(* IEC 61131-3 sources: Jacob-Formschaumtechnik-ISEL-CNC-Retrofit/twincat/PLC/src/0_Main, 9 files *)

(* ---- GVL_AlarmCatalog.st ---- *)
(* Meldekatalog, einzige Quelle fuer ID und Klasse je Slot (Befund 11). Slot-Nummer = Index in aCond,
   siehe E_AlarmSlot. Klassen: 0 Info, 1 Warnung, 2 Vorschubhalt, 3 Abbruch, 4 Antriebe aus.
   Slot 12 (Referenzverlust) ist R1, Slot 13 (HMI-Verbindung) R2. Texte pflegt die HMI-Seite. *)
VAR_GLOBAL CONSTANT
    aAlarmId    : ARRAY[0..14] OF INT := [100, 101, 110, 120, 200, 201, 202, 203, 300, 301, 302, 310, 320, 330, 900];
    (* Befund 15: 200 (FU-Stoerung) und 302 (Endschalter) sind R3 statt R4. Die Achsregler bleiben an,
       das Programm wird abgebrochen, vom Endschalter kann in Hand freigefahren werden. [Annahme, mit Kunde abstimmen] *)
    aAlarmClass : ARRAY[0..14] OF INT := [4, 3, 3, 2, 3, 3, 3, 1, 4, 4, 3, 4, 1, 2, 4];
END_VAR

(* ---- GVL_Config.st ---- *)
(* Build-Konfiguration (Befund 9). Die Antriebsabbildung wird hier gewaehlt. Solange nur das
   Simulationsabbild fertig ist, laeuft die Maschine nur damit. Fuer jede andere Variante bleibt die
   Maschine gesperrt (FB_AxisMap_Canopen meldet Fehler FFFF0001), bis die echte Abbildung existiert.
   Auf einer realen Maschine darf bSimulationBuild nicht TRUE sein. *)
VAR_GLOBAL CONSTANT
    eDriveVariant   : E_DriveVariant := E_DriveVariant.Simulation;
    bSimulationBuild: BOOL := (eDriveVariant = E_DriveVariant.Simulation);   (* G-06: nie getrennt von der Antriebsvariante setzen *)
    sSwVersion      : STRING(15) := '0.12.0';   (* G-18: bei jedem Tag mitpflegen, auch in FB_ParamInit *)
    (* Befund 20: Maschinenkennung kommt aus GVL_Persistent.nMachineId, nicht aus dem Code.
       Nur im Simulationsbuild gilt bei nicht gesetzter Kennung (0) die Kennung 1 [Annahme]. *)
    nMachineIdSimDefault : UINT := 1;
    (* Achsnummerierung zentral (Befund 16). HMI- und CNC-Achse: 1 = X, 2 = Y, 3 = Z [Annahme CNC-Kanal].
       Referenzgruppe: 1 = Z, 2 = X, 3 = Y. Antrieb: 1 = Y1, 2 = Y2, 3 = X, 4 = Z [Annahme]. *)
    aHmiAxisToGroup  : ARRAY[1..3] OF USINT := [2, 3, 1];
    aGroupToHmiAxis  : ARRAY[1..3] OF USINT := [3, 1, 2];
    aDriveToHmiAxis  : ARRAY[1..4] OF USINT := [2, 2, 1, 3];
    aDriveToGroup    : ARRAY[1..4] OF USINT := [3, 3, 2, 1];
    (* Befund 15: Verzoegerung der Reglerabschaltung bei R4, damit die CNC gefuehrt bremst [Annahme] *)
    tR4DriveOffDelay : TIME := T#500MS;
END_VAR

(* ---- GVL_HMI.st ---- *)
VAR_GLOBAL
    stCmd : ST_HmiCmd;     (* HMI -> SPS *)
    stSts : ST_HmiSts;     (* SPS -> HMI *)
    stJournal : ST_HmiJournal;  (* SPS -> HMI, Meldejournal (Befund 21), Kopie von GVL_Persistent.stJournal *)
END_VAR

(* ---- GVL_HmiCnc.st ---- *)
VAR_GLOBAL
    stCncSts : ST_HmiCncSts;     (* SPS -> HMI *)
    stCncCmd : ST_HmiCncCmd;     (* HMI -> SPS *)
END_VAR

(* ---- GVL_IO.st ---- *)
(* Prozessabbild der Maschine. Die Verknuepfung mit den Klemmen erfolgt erst nach
   Klemmenwahl und Schaltplan, bis dahin gibt es hier nur Variablen ohne Adresse (Simulation).
   Ruhestrom: FALSE = Fehler/ausgeloest bei allen Sicherheits- und Endschaltersignalen. *)
VAR_GLOBAL
    (* Eingaenge *)
    bSafetyRelayFeedback : BOOL;   (* Pilz-Relais Rueckmeldung *)
    bDoorClosed          : BOOL;
    bAirOk               : BOOL;
    bExtractionOk        : BOOL;
    bFuReady             : BOOL;   (* Commander SK bereit *)
    bFuAtSpeed           : BOOL;   (* [Annahme] Drehzahl erreicht *)
    bSpindlePtcOk        : BOOL;
    bKeyAuto             : BOOL;   (* [offen] nur falls Schluesselschalter vorhanden *)
    bFieldbusOk          : BOOL;   (* EtherCAT/CANopen Status *)
    (* Ausgaenge *)
    bSpindleRun          : BOOL;
    bSpindleCcw          : BOOL;
    rSpindleVolt         : REAL;   (* EL4002 Kanal 1, 0..10 V *)
    bExtractionOut       : BOOL;
    bBlowAirOut          : BOOL;
    bVacuumOut           : BOOL;
    (* Achsen, vier Stueck: 1=Y1 Portal links, 2=Y2 Portal rechts, 3=X Quer, 4=Z [Annahme] *)
    aAxis                : ARRAY[1..4] OF ST_AxisDrive;
    (* Einspeisung fuer Simulation und Test (wirkt nur im Simulationsabbild FB_AxisMap_Simulation) *)
    aSimLimitPlus  : ARRAY[1..4] OF BOOL;
    aSimLimitMinus : ARRAY[1..4] OF BOOL;
    aSimFault      : ARRAY[1..4] OF BOOL;
END_VAR

(* ---- GVL_Machine.st ---- *)
(* Zustandsgroessen und CNC-Schnittstelle (Signale aus/zur CNC kommen spaeter ueber Tc2_CncHli). *)
VAR_GLOBAL
    stParams       : ST_MachineParams;
    bParamsLoaded  : BOOL;
    (* von der CNC [offen, HLI-Anbindung folgt] *)
    nCncMCode      : INT;
    bCncMStrobe    : BOOL;
    nCncToolNo     : UINT;
    bCncProgramDone: BOOL;
    bCncProgramActive : BOOL;  (* Programm laeuft oder Achsen fahren noch (Befund 4) *)
    rCncSpindleRpm : REAL;     (* S-Wert aus dem NC-Programm, 1/min (Befund 10) *)
    aCncHomed      : ARRAY[1..3] OF BOOL;
    (* zur CNC *)
    bCncStartReq   : BOOL;
    bCncHoldReq    : BOOL;
    bCncAbortReq   : BOOL;
    bCncMAck       : BOOL;
    bCncJogPlus    : BOOL;
    bCncJogMinus   : BOOL;
    nCncJogAxis    : USINT;
    bCncJogRapid   : BOOL;
    bCncHomeReq    : BOOL;
    nCncHomeGroup  : USINT;
    bCncSingleBlock: BOOL;
    bCncDryRun     : BOOL;
    bCncOptStop    : BOOL;
    rCncJogStepMm  : REAL;
    bCncHandwheel  : BOOL;
    nCncHandwheelAxis  : USINT;
    nCncHandwheelRatio : USINT;
    bHasHandwheel  : BOOL;     (* [offen] nur M1 mit Bestandsgeraet *)
    bCncJogCreep   : BOOL;     (* Freifahren vom Endschalter: CNC soll im Schleichgang tippen (HLI-Anbindung offen) *)
END_VAR

(* ---- GVL_Persistent.st ---- *)
{attribute 'qualified_only'}
(* Persistente Daten (Befunde 20 und 21). Ueberleben Neustart und Online-Change.
   nMachineId ist die Maschinenkennung des Geraets, gesetzt bei der Inbetriebnahme (0 = nicht gesetzt,
   Maschine bleibt gesperrt, Meldung 900). Damit laeuft ein Softwarestand auf allen Maschinen (LH-2.11.4).
   [offen] Schreibweg ueber die Service-Seite der HMI, bis dahin per ADS. *)
VAR_GLOBAL PERSISTENT
    nMachineId    : UINT;
    nOperatingSec : UDINT;            (* Betriebssekunden *)
    nSpindleSec   : UDINT;            (* Spindellaufzeit in Sekunden *)
    stJournal     : ST_HmiJournal;    (* Meldejournal *)
END_VAR

(* ---- PRG_Main.st ---- *)
(* Hauptprogramm. Aufrufreihenfolge fest: Eingaenge -> Sicherheit -> Achsen -> Meldungen ->
   Verriegelungen -> Zustand -> Geraete -> HMI-Status. Rueckwirkungen zwischen den Bausteinen
   laufen bewusst mit einem Zyklus Verzoegerung, damit keine Schleifen entstehen. *)
PROGRAM PRG_Main
VAR
    fbParamInit: FB_ParamInit;
    fbCncMirror: FB_CncMirror;
    fbParam    : FB_ParamCheck;
    aGrpOfAxis : ARRAY[1..4] OF INT := [3, 3, 2, 1];   (* Achse 1,2 (Y1,Y2) = Gruppe 3, Achse 3 (X) = Gruppe 2, Achse 4 (Z) = Gruppe 1 *)
    fbSafety   : FB_SafetyMonitor;
    fbAxisSim  : ARRAY[1..4] OF FB_AxisMap_Simulation;
    fbSupervisor : FB_AxisSupervisor;
    fbAlarms   : FB_AlarmList;
    fbJournal  : FB_AlarmJournal;
    fbInterlocks : FB_Interlocks;
    fbState    : FB_MachineState;
    fbMode     : FB_OpModeManager;
    fbSpindle  : FB_Spindle;
    fbMFunc    : FB_MFunctions;
    fbTool     : FB_ToolChange;
    fbHoming   : FB_Homing;
    fbJog      : FB_Jog;
    aCond      : ARRAY[0..14] OF BOOL;
    aHomeReq   : ARRAY[1..3] OF BOOL;
    fbAxisCan  : ARRAY[1..4] OF FB_AxisMap_Canopen;
    tonExtraction : TON;
    i          : INT;
    bStandstill: BOOL;
    bSimulation: BOOL := TRUE;     (* bis die Hardwareabbildung steht, immer Simulation *)
    nVersionDummy : INT;
    tonUptime  : TON;
    tonSpindleUptime : TON;
    dwSecTick  : UDINT;
    dtNow      : DT;
    nMachineIdEff : UINT;     (* wirksame Maschinenkennung (Befund 20) *)
    nSysTime   : ULINT;       (* UTC, 100 ns seit 1.1.1601 *)
    bLimitFreeRun : BOOL;     (* Freifahren vom Endschalter erlaubt (Befund 15) *)
    bOtherR3   : BOOL;
    nCls       : INT;
    bHandSpindleBlock : BOOL; (* Hand-Spindel gesperrt bis bSpindleOn einmal FALSE war (Lebenszeichen weg, nicht Hand) *)
    bHandSpindleOn : BOOL;    (* wirksame Hand-Anforderung Spindel *)
    tofModeBlocked : TOF;     (* Hinweis "Betriebsartwechsel abgelehnt" fuer die HMI halten *)
    bLimHitPlus      : BOOL;
    bLimHitMinus     : BOOL;
    bJogPlusBlocked  : BOOL;
    bJogMinusBlocked : BOOL;
    rtHandOn         : R_TRIG;
    bHandCcw         : BOOL;
    bDryRunEff       : BOOL;
    bSpindleLocked   : BOOL;
    bVacuumReq       : BOOL;
    bHomingLostInRun : BOOL;
    bToolChangeDoor  : BOOL;
END_VAR

(* 1. Parameter: initialisieren und pruefen, bei unplausiblen Werten bleibt die Maschine gesperrt *)
(* Befund 20: Kennung aus dem Geraet (persistent), nur im Simulationsbuild Ersatzwert bei 0 *)
nMachineIdEff := GVL_Persistent.nMachineId;
IF nMachineIdEff = 0 AND GVL_Config.bSimulationBuild THEN nMachineIdEff := GVL_Config.nMachineIdSimDefault; END_IF
fbParamInit(nMachineId := nMachineIdEff, stParams := GVL_Machine.stParams);
GVL_Machine.bParamsLoaded := fbParamInit.bLoaded;
fbParam(nIdExpected := nMachineIdEff, nIdLoaded := GVL_Machine.stParams.nMachineId,
        sVerExpected := GVL_Machine.stParams.sSwVersionExpected, sVerRunning := GVL_Config.sSwVersion,
        bParamsLoaded := GVL_Machine.bParamsLoaded);

(* 2. Sicherheit *)
fbSafety(bRelayFeedbackOk := GVL_IO.bSafetyRelayFeedback, bDoorClosed := GVL_IO.bDoorClosed,
         bFieldbusOk := GVL_IO.bFieldbusOk, bAck := GVL_HMI.stCmd.bAck, bAirOk := GVL_IO.bAirOk);

(* 3. Achsen *)
FOR i := 1 TO 4 DO
    GVL_IO.aAxis[i].bEnableReq := fbState.bEnableDrives;
    GVL_IO.aAxis[i].bResetReq  := GVL_HMI.stCmd.bAck;     (* Antriebsfehler quittieren (Befund 14) *)
    IF GVL_Config.eDriveVariant = E_DriveVariant.Simulation THEN
    fbAxisSim[i](bSafeEnable := fbSafety.bDrivesAllowed,
                 bHomeReset := fbHoming.aResetHomed[GVL_Config.aDriveToGroup[i]],
                 bHomeCmd := fbHoming.bHomeCmd AND fbHoming.nActiveGroup = GVL_Config.aDriveToGroup[i],
                 bInjLimitPlus := GVL_IO.aSimLimitPlus[i], bInjLimitMinus := GVL_IO.aSimLimitMinus[i],
                 bInjFault := GVL_IO.aSimFault[i],
                 stAxis := GVL_IO.aAxis[i]);
    ELSE
        (* Befund 9: echte Abbildung fehlt, FB_AxisMap_Canopen sperrt die Maschine (Fehler FFFF0001) *)
        fbAxisCan[i](bSafeEnable := fbSafety.bDrivesAllowed, stAxis := GVL_IO.aAxis[i]);
    END_IF
END_FOR
(* Einheitlicher Referenzstatus (Befund 3): einzige Quelle ist GVL_IO.aAxis[].bHomed.
   Gruppen 1 = Z, 2 = X, 3 = Y (beide Portalseiten). *)
GVL_Machine.aCncHomed[1] := GVL_IO.aAxis[4].bHomed;
GVL_Machine.aCncHomed[2] := GVL_IO.aAxis[3].bHomed;
GVL_Machine.aCncHomed[3] := GVL_IO.aAxis[1].bHomed AND GVL_IO.aAxis[2].bHomed;
GVL_HmiCnc.stCncSts.aAxis[1].bHomed := GVL_Machine.aCncHomed[2];   (* HMI-Achse 1 = X *)
GVL_HmiCnc.stCncSts.aAxis[2].bHomed := GVL_Machine.aCncHomed[3];   (* HMI-Achse 2 = Y *)
GVL_HmiCnc.stCncSts.aAxis[3].bHomed := GVL_Machine.aCncHomed[1];   (* HMI-Achse 3 = Z *)
fbSupervisor(bEnableCmd := fbState.bEnableDrives, bFieldbusOk := GVL_IO.bFieldbusOk,
             bHomingActive := fbHoming.bBusy, rMaxFollowErr := 1.0, aAxis := GVL_IO.aAxis);
bStandstill := fbSpindle.bStandstillOk AND fbState.eState <> E_MachState.Execute AND NOT fbJog.bJogPlusReq AND NOT fbJog.bJogMinusReq;

(* 4. Meldungen *)
(* Werkzeugwechsel mit Tuerfreigabe: Tuer offen und Spindel steht. Dann sind Tuer-Meldung und das dadurch abfallende
   Sicherheitsrelais kein Abbruchgrund, das Programm bleibt gehalten. Sonst ist eine offene Tuer weiter ein Abbruch. *)
bToolChangeDoor := fbTool.bDoorRelease AND NOT GVL_IO.bDoorClosed AND GVL_IO.bFieldbusOk;
aCond[0]  := NOT GVL_IO.bSafetyRelayFeedback AND NOT bToolChangeDoor;
aCond[1]  := NOT GVL_IO.bDoorClosed AND NOT bToolChangeDoor;
aCond[2]  := GVL_Machine.stParams.bAirMonitoring AND NOT GVL_IO.bAirOk;
(* Absaugung: Rueckmeldung darf nach dem Einschalten tFeedbackTimeout dauern (Befund 12) *)
tonExtraction(IN := NOT GVL_IO.bExtractionOk AND GVL_IO.bExtractionOut, PT := GVL_Machine.stParams.tFeedbackTimeout);
aCond[3]  := tonExtraction.Q;
aCond[4]  := NOT GVL_IO.bFuReady;
aCond[5]  := fbSpindle.bPtcTrip;
aCond[6]  := fbSpindle.bNoFeedback;
aCond[7]  := fbSpindle.bLockedSetup;
aCond[8]  := fbSupervisor.bAnyFault OR fbSupervisor.bEnableTimeout;
aCond[9]  := fbSupervisor.bFollowErr;
aCond[10] := fbSupervisor.bAnyHwLimit;
aCond[11] := NOT GVL_IO.bFieldbusOk;
aCond[12] := fbSupervisor.bHomingLost;
aCond[13] := NOT fbJog.bHmiLinkOk;
aCond[14] := fbParam.bMismatch;
fbAlarms(aCond := aCond, bAck := GVL_HMI.stCmd.bAck);
(* Befund 21: Zeitstempel UTC, Journal persistent, HMI liest die Kopie *)
nSysTime := F_GetSystemTime();
IF nSysTime > 116444736000000000 THEN
    dtNow := DWORD_TO_DT(ULINT_TO_DWORD((nSysTime - 116444736000000000) / 10000000));
END_IF
fbJournal(aCond := aCond, aId := GVL_AlarmCatalog.aAlarmId, aClass := GVL_AlarmCatalog.aAlarmClass,
          dtNow := dtNow, stJournal := GVL_Persistent.stJournal);
GVL_HMI.stJournal := GVL_Persistent.stJournal;

(* Befund 15: Steht nur der Endschalter (302, R3) an, darf in Hand im Schleichgang freigefahren werden.
   [offen] Richtungssperre zur Endschalterseite liegt in CNC/Antrieb (Softwareendlage, Endschalterlogik). *)
bOtherR3 := FALSE;
FOR i := 0 TO 14 DO
    nCls := GVL_AlarmCatalog.aAlarmClass[i];
    IF i <> 10 (* E_AlarmSlot.HwLimitHit *) AND nCls >= 3 AND (fbAlarms.aList[i].bActive OR fbAlarms.aList[i].bLatched) THEN
        bOtherR3 := TRUE;
    END_IF
END_FOR
bLimitFreeRun := aCond[10] AND NOT bOtherR3;   (* Slot 10 = E_AlarmSlot.HwLimitHit *)

(* 5. Betriebsart und Verriegelungen *)
(* Befund 17: Wechsel nur im echten Stillstand, ohne Referenzfahrt und ohne offene Werkzeugwechsel-Aufforderung *)
fbMode(eRequest := GVL_HMI.stCmd.eModeRequest,
       bStandstill := bStandstill AND fbInterlocks.bModeChangeOk AND NOT fbHoming.bBusy AND NOT fbTool.bRequest,
       bHasKeySwitch := FALSE, bKeyAuto := GVL_IO.bKeyAuto);
(* Abgelehnter Wunsch wird verworfen, sonst fuehrte die SPS ihn beim naechsten Stillstand verspaetet aus.
   Der Hinweis bleibt 3 s fuer die HMI stehen. *)
IF fbMode.bChangeBlocked THEN
    GVL_HMI.stCmd.eModeRequest := fbMode.eMode;
END_IF
tofModeBlocked(IN := fbMode.bChangeBlocked, PT := T#3S);
fbInterlocks(eMode := fbMode.eMode, eState := fbState.eState, bSafetyOk := fbSafety.bSafetyOk,
             bAllHomed := fbSupervisor.bAllHomed, bDrivesEnabled := fbSupervisor.bAllEnabled,
             bHmiLinkOk := fbJog.bHmiLinkOk, bAnyR2OrHigher := fbAlarms.bAnyR2OrHigher,
             bAnyR3OrHigher := fbAlarms.bAnyR3OrHigher, bAirOk := GVL_IO.bAirOk OR NOT GVL_Machine.stParams.bAirMonitoring,
             bHomingBusy := fbHoming.bBusy, bLimitFreeRun := bLimitFreeRun);

(* 6. Zustand *)
(* G-10: Geht die Referenz im laufenden oder gehaltenen Programm verloren, wirkt das wie R3 (Abbruch). Sonst nur Warnung R1. *)
bHomingLostInRun := fbSupervisor.bHomingLost AND (fbState.eState = E_MachState.Execute OR fbState.eState = E_MachState.Held);
fbState(bSafetyOk := fbSafety.bSafetyOk, bDrivesAllowed := fbSafety.bDrivesAllowed,
        bAnyR2OrHigher := fbAlarms.bAnyR2OrHigher OR bHomingLostInRun,
        bAnyR3OrHigher := fbAlarms.bAnyR3OrHigher OR bHomingLostInRun,
        bAnyR4 := fbAlarms.bAnyR4, bAckPending := fbAlarms.bAckPending,
        bStartOk := fbInterlocks.bProgramStartOk AND NOT fbTool.bHoldProgram,
        bStartCmd := GVL_HMI.stCmd.bStart, bHoldCmd := GVL_HMI.stCmd.bHold OR fbMFunc.bProgramHalt,
        bAbortCmd := GVL_HMI.stCmd.bAbort, bProgramDone := GVL_Machine.bCncProgramDone,
        bProgramActive := GVL_Machine.bCncProgramActive,
        bAck := GVL_HMI.stCmd.bAck, tR4OffDelay := GVL_Config.tR4DriveOffDelay,
        bDoorOpenAllowed := bToolChangeDoor);

(* 7. Geraete: Spindel (M3/M4 aus Programm, in Hand von der HMI) *)
(* Hand-Spindel: Nach Lebenszeichenverlust oder ausserhalb Hand setzt die SPS bSpindleOn zurueck und sperrt,
   bis bSpindleOn FALSE gesehen wurde. Ein stehender Pegel startet die Spindel so nie von selbst wieder. *)
IF NOT fbJog.bHmiLinkOk OR fbMode.eMode <> E_OpMode.Hand THEN
    bHandSpindleBlock := TRUE;
    GVL_HMI.stCmd.bSpindleOn := FALSE;
ELSIF NOT GVL_HMI.stCmd.bSpindleOn THEN
    bHandSpindleBlock := FALSE;
END_IF
bHandSpindleOn := GVL_HMI.stCmd.bSpindleOn AND NOT bHandSpindleBlock;
(* G-11: Drehrichtung wird beim Einschalten festgehalten, Umschalten bei laufender oder wartender Spindel startet nichts *)
rtHandOn(CLK := bHandSpindleOn);
IF rtHandOn.Q THEN bHandCcw := GVL_HMI.stCmd.bSpindleCcw; END_IF
(* G-12: Trockenlauf wirkt nur in Auto und nur so, wie er beim Programmstart stand (nicht mitten im Programm) *)
IF fbState.eState <> E_MachState.Execute AND fbState.eState <> E_MachState.Held THEN
    bDryRunEff := GVL_HMI.stCmd.bDryRun;
END_IF
bSpindleLocked := fbMode.eMode = E_OpMode.Setup OR (fbMode.eMode = E_OpMode.Auto AND bDryRunEff);
fbMFunc(nMCode := GVL_Machine.nCncMCode, bMStrobe := GVL_Machine.bCncMStrobe,
        bSpindleOk := fbInterlocks.bSpindleOk, bAuxOk := fbInterlocks.bAuxOk,
        bReset := fbState.bSpindleStop OR GVL_Machine.bCncProgramDone, bOptStop := GVL_HMI.stCmd.bOptStop,
        bSpindleRunning := fbSpindle.bRunning, bSpindleSkip := bSpindleLocked);
fbSpindle(bRelease := fbInterlocks.bSpindleOk AND NOT fbState.bSpindleStop AND NOT fbTool.bSpindleLock,
          bStop := fbState.bSpindleStop,
          bSetupLocked := bSpindleLocked,
          bAllowPend := fbMode.eMode = E_OpMode.Auto,   (* G-11: nur das Programm darf auf Stillstand warten, Hand-Start wird sonst verworfen *)
          bStartCw := (fbMFunc.bSpindleCw AND fbMode.eMode = E_OpMode.Auto) OR (bHandSpindleOn AND NOT bHandCcw),
          bStartCcw := (fbMFunc.bSpindleCcw AND fbMode.eMode = E_OpMode.Auto) OR (bHandSpindleOn AND bHandCcw),
          rSetRpm := SEL(fbMode.eMode = E_OpMode.Auto, GVL_HMI.stCmd.rSpindleSetRpm, GVL_Machine.rCncSpindleRpm),
          rOverridePct := UINT_TO_REAL(GVL_HmiCnc.stCncSts.nOvrSpindle),
          bFuReady := GVL_IO.bFuReady, bFuAtSpeed := GVL_IO.bFuAtSpeed, bPtcOk := GVL_IO.bSpindlePtcOk,
          bAckReset := GVL_HMI.stCmd.bAck, rMaxRpm := GVL_Machine.stParams.rSpindleMaxRpm,
          rMinRpm := GVL_Machine.stParams.rSpindleMinRpm, rVoltMax := GVL_Machine.stParams.rSpindleVoltMax,
          tRunUp := GVL_Machine.stParams.tSpindleRunUp, tStandstill := GVL_Machine.stParams.tSpindleStandstill);
GVL_IO.bSpindleRun  := fbSpindle.bRunCmd;
GVL_IO.bSpindleCcw  := fbSpindle.bDirCcw;
GVL_IO.rSpindleVolt := fbSpindle.rVoltOut;

fbTool(bM6Request := fbMFunc.bToolChangeReq, nToolNo := GVL_Machine.nCncToolNo,
       bSpindleStopped := fbSpindle.bStandstillOk, bConfirm := GVL_HMI.stCmd.bToolChangeDone,
       bAbort := GVL_HMI.stCmd.bAbort OR fbState.eState = E_MachState.EStop OR fbState.eState = E_MachState.Aborted
                 OR fbState.eState = E_MachState.Fault);   (* G-05: Anforderung faellt bei Abbruch, R3 und NOT-HALT *)

(* Hilfsausgaenge: von Hand oder per M-Code, nur mit Freigabe *)
GVL_IO.bExtractionOut := fbInterlocks.bAuxOk AND (fbMFunc.bExtraction OR GVL_HMI.stCmd.bExtraction);
GVL_IO.bBlowAirOut    := fbInterlocks.bAuxOk AND (fbMFunc.bBlowAir OR GVL_HMI.stCmd.bBlowAir);
(* G-04: Vakuum (Werkstueckspannung) bleibt bei Abbruch und NOT-HALT gehalten. Einschalten nur mit Freigabe. *)
bVacuumReq := fbMFunc.bVacuum OR GVL_HMI.stCmd.bVacuum;
GVL_IO.bVacuumOut     := bVacuumReq AND (fbInterlocks.bAuxOk OR GVL_IO.bVacuumOut);

(* 8. Referenzieren und Tippen *)
(* Zuordnung HMI-Achse (1=X, 2=Y, 3=Z) zu Referenzgruppe (1=Z, 2=X, 3=Y) *)
aHomeReq[1] := GVL_HMI.stCmd.bHomeAxis[3];
aHomeReq[2] := GVL_HMI.stCmd.bHomeAxis[1];
aHomeReq[3] := GVL_HMI.stCmd.bHomeAxis[2];
fbHoming(bStart := GVL_HMI.stCmd.bHomeRequest, aStartAxis := aHomeReq,
         bAbort := GVL_HMI.stCmd.bAbort OR GVL_HMI.stCmd.bHomeAbort,
         bHomingOk := fbInterlocks.bHomingOk, aHomed := GVL_Machine.aCncHomed);
(* G-01: Endschalter je Seite der gewaehlten Achse (HMI 1=X -> Antrieb 3, 2=Y -> Antriebe 1 und 2, 3=Z -> Antrieb 4).
   Ruhestrom: FALSE = ausgeloest. [Annahme] Tippen+ faehrt zur Plus-Seite. Ist ein Endschalter ausgeloest, ist Tippen
   nur fuer die betroffene Achse und nur in Gegenrichtung erlaubt, ohne Eilgang. *)
bLimHitPlus := FALSE; bLimHitMinus := FALSE;
CASE GVL_HMI.stCmd.nJogAxis OF
    1: bLimHitPlus  := NOT GVL_IO.aAxis[3].bHwLimitPlus;
       bLimHitMinus := NOT GVL_IO.aAxis[3].bHwLimitMinus;
    2: bLimHitPlus  := NOT GVL_IO.aAxis[1].bHwLimitPlus  OR NOT GVL_IO.aAxis[2].bHwLimitPlus;
       bLimHitMinus := NOT GVL_IO.aAxis[1].bHwLimitMinus OR NOT GVL_IO.aAxis[2].bHwLimitMinus;
    3: bLimHitPlus  := NOT GVL_IO.aAxis[4].bHwLimitPlus;
       bLimHitMinus := NOT GVL_IO.aAxis[4].bHwLimitMinus;
END_CASE
bJogPlusBlocked  := bLimHitPlus;
bJogMinusBlocked := bLimHitMinus;
IF aCond[10] AND NOT (bLimHitPlus OR bLimHitMinus) THEN
    bJogPlusBlocked := TRUE; bJogMinusBlocked := TRUE;   (* Endschalter an einer anderen Achse: diese Achse bleibt stehen *)
END_IF
GVL_Machine.bCncJogCreep := bLimitFreeRun;   (* CNC: Freifahren nur im Schleichgang (HLI-Anbindung offen) *)
fbJog(bJogOk := fbInterlocks.bJogOk, bPlus := GVL_HMI.stCmd.bJogPlus, bMinus := GVL_HMI.stCmd.bJogMinus,
      bPlusBlocked := bJogPlusBlocked, bMinusBlocked := bJogMinusBlocked,
      nAxis := GVL_HMI.stCmd.nJogAxis, bRapid := GVL_HMI.stCmd.bJogRapid AND NOT bLimitFreeRun AND GVL_HmiCnc.stCncSts.nSpeedLimitActivePct >= 50,
      nHeartbeat := GVL_HMI.stCmd.nHeartbeat, tHmiTimeout := GVL_Machine.stParams.tHmiTimeout);

(* CNC-Spiegel (Simulation, bis TF5200 verfuegbar ist) *)
fbCncMirror(bStandstill := fbState.eState <> E_MachState.Execute AND fbState.eState <> E_MachState.Held
                           AND NOT GVL_Machine.bCncProgramActive,
            stCmd := GVL_HmiCnc.stCncCmd, stSts := GVL_HmiCnc.stCncSts);

(* 9. Anforderungen an die CNC *)
GVL_Machine.bCncStartReq := fbState.bCncStart;
GVL_Machine.bCncHoldReq  := fbState.bCncHold OR fbTool.bHoldProgram;
GVL_Machine.bCncAbortReq := fbState.bCncAbort;
GVL_Machine.bCncMAck     := fbMFunc.bAck;
GVL_Machine.bCncJogPlus  := fbJog.bJogPlusReq;
GVL_Machine.bCncJogMinus := fbJog.bJogMinusReq;
GVL_Machine.nCncJogAxis  := fbJog.nAxisReq;
GVL_Machine.bCncJogRapid := fbJog.bRapidReq;
GVL_Machine.bCncHomeReq  := fbHoming.bHomeCmd;
GVL_Machine.nCncHomeGroup:= fbHoming.nActiveGroup;
GVL_Machine.bCncSingleBlock := GVL_HMI.stCmd.bSingleBlock;
GVL_Machine.bCncDryRun   := bDryRunEff AND fbMode.eMode = E_OpMode.Auto;
GVL_Machine.bCncOptStop  := GVL_HMI.stCmd.bOptStop;
GVL_Machine.rCncJogStepMm := GVL_HMI.stCmd.rJogStepMm;
(* Handrad: nur freigegeben, wenn vorhanden, in Hand und Tippen erlaubt *)
GVL_Machine.bCncHandwheel := GVL_Machine.bHasHandwheel AND GVL_HMI.stCmd.bHandwheelEnable AND fbInterlocks.bJogOk;
GVL_Machine.nCncHandwheelAxis  := GVL_HMI.stCmd.nHandwheelAxis;
GVL_Machine.nCncHandwheelRatio := GVL_HMI.stCmd.nHandwheelRatio;

(* 10. Status an die HMI *)
(* Befund 21: Betriebs- und Spindellaufzeit persistent, Sekundentakt *)
tonUptime(IN := TRUE, PT := T#1S);
IF tonUptime.Q THEN
    dwSecTick := dwSecTick + 1;
    GVL_Persistent.nOperatingSec := GVL_Persistent.nOperatingSec + 1;
    IF fbSpindle.bRunCmd THEN GVL_Persistent.nSpindleSec := GVL_Persistent.nSpindleSec + 1; END_IF
    tonUptime(IN := FALSE);
END_IF
GVL_HMI.stSts.eMode          := fbMode.eMode;
GVL_HMI.stSts.eState         := fbState.eState;
GVL_HMI.stSts.bSafetyOk      := fbSafety.bSafetyOk;
GVL_HMI.stSts.bDrivesEnabled := fbSupervisor.bAllEnabled;
GVL_HMI.stSts.bAllHomed      := fbSupervisor.bAllHomed;
GVL_HMI.stSts.bHmiLinkOk     := fbJog.bHmiLinkOk;
GVL_HMI.stSts.bSpindleRunning:= fbSpindle.bRunning;
GVL_HMI.stSts.rSpindleActRpm := SEL(fbSpindle.bRunning, 0.0, fbSpindle.rActRpm);   (* Sollwert nur bei Drehzahl erreicht anzeigen (Befund 13) *)
GVL_HMI.stSts.bExtractionOn  := GVL_IO.bExtractionOut;
GVL_HMI.stSts.bBlowAirOn     := GVL_IO.bBlowAirOut;
GVL_HMI.stSts.bVacuumOn      := GVL_IO.bVacuumOut;
GVL_HMI.stSts.bToolChangeReq := fbTool.bRequest;
GVL_HMI.stSts.nToolChangeNo  := fbTool.nRequestedTool;
GVL_HMI.stSts.nTopAlarmId    := fbAlarms.nTopId;
GVL_HMI.stSts.eTopAlarmClass := F_ToFaultClass(fbAlarms.nTopClass);
GVL_HMI.stSts.nActiveAlarms  := fbAlarms.nActive;
GVL_HMI.stSts.nMachineId     := GVL_Machine.stParams.nMachineId;
GVL_HMI.stSts.sSwVersion     := GVL_Config.sSwVersion;
GVL_HMI.stSts.bSimulationActive := GVL_Config.bSimulationBuild;
GVL_HMI.stSts.bModeChangeBlocked := tofModeBlocked.Q;
GVL_HMI.stSts.dwOperatingSec := GVL_Persistent.nOperatingSec;
GVL_HMI.stSts.dwSpindleSec   := GVL_Persistent.nSpindleSec;
GVL_HMI.stSts.nHeartbeatEcho := GVL_HMI.stCmd.nHeartbeat;
GVL_HMI.stSts.bLimitFreeRun  := bLimitFreeRun;
GVL_HMI.stSts.bToolChangeDoorRelease := fbTool.bDoorRelease;
GVL_HMI.stSts.bHandwheelActive := GVL_Machine.bCncHandwheel;
GVL_HMI.stSts.eHomeState[1]  := fbHoming.eHomeState[2];   (* X *)
GVL_HMI.stSts.eHomeState[2]  := fbHoming.eHomeState[3];   (* Y *)
GVL_HMI.stSts.eHomeState[3]  := fbHoming.eHomeState[1];   (* Z *)
GVL_HMI.stSts.nHomeStep      := fbHoming.nStepOut;
GVL_HMI.stSts.aAlarms        := fbAlarms.aList;
GVL_HMI.stSts.aDrive         := GVL_IO.aAxis;
GVL_HMI.stSts.bFieldbusOk    := GVL_IO.bFieldbusOk;
GVL_HMI.stSts.bFuFault       := NOT GVL_IO.bFuReady;
GVL_HMI.stSts.bPtcTrip       := fbSpindle.bPtcTrip;

(* 11. Befund 16: Impulse aus der HMI loescht die SPS nach der Auswertung in diesem Zyklus.
   Die HMI setzt nur TRUE (Einzelfeld schreiben, nicht die ganze Struktur), ein Impuls geht so nie verloren. *)
GVL_HMI.stCmd.bStart          := FALSE;
GVL_HMI.stCmd.bHold           := FALSE;
GVL_HMI.stCmd.bAbort          := FALSE;
GVL_HMI.stCmd.bAck            := FALSE;
GVL_HMI.stCmd.bHomeRequest    := FALSE;
GVL_HMI.stCmd.bHomeAbort      := FALSE;
GVL_HMI.stCmd.bToolChangeDone := FALSE;
GVL_HMI.stCmd.bHomeAxis[1]    := FALSE;
GVL_HMI.stCmd.bHomeAxis[2]    := FALSE;
GVL_HMI.stCmd.bHomeAxis[3]    := FALSE;
GVL_HmiCnc.stCncCmd.bProgramLoad   := FALSE;
GVL_HmiCnc.stCncCmd.bTableWrite    := FALSE;
GVL_HmiCnc.stCncCmd.bWcsSetCurrent := FALSE;
END_PROGRAM

(* ---- PRG_Test.st ---- *)
(* Simulationstest der Grundfunktionen (nur im Simulations-Build, GVL_Config.bSimulationBuild).
   Starten: bTestEnable online auf TRUE setzen. Der Test speist Eingaenge und HMI-Kommandos ein und prueft
   Referenz, Tippen, NOT-HALT und Spindel gegen die Fehlerfaelle aus dem Gutachten (kein Selbstanlauf nach
   Quittierung). Ergebnis: bTestDone, nFails, sFirstFail. Rueckgabe in der Runtime lesen. *)
PROGRAM PRG_Test
VAR
    bTestEnable : BOOL;                 (* online auf TRUE setzen *)
    bTestDone   : BOOL;
    nFails      : INT;
    sFirstFail  : STRING(100);
    nStep       : INT;
    tWait       : TIME;
    tonStep     : TON;
    tonHb       : TON;
    bNext       : BOOL;
    bRelay      : BOOL := TRUE;         (* Rueckmeldung Sicherheitsrelais, NOT-HALT = FALSE *)
    bFailNow    : BOOL;
    sMsg        : STRING(100);
    bHbStop     : BOOL;                 (* TRUE = simuliertes Lebenszeichen der HMI ausgefallen *)
    nIdx        : INT;
    bDoor       : BOOL := TRUE;         (* Tuer geschlossen *)
END_VAR

(* G-06: Der Test schreibt Sicherheitseingaenge und darf nur mit dem Simulationsabbild laufen *)
IF NOT (bTestEnable AND GVL_Config.bSimulationBuild AND GVL_Config.eDriveVariant = E_DriveVariant.Simulation) THEN
    bHbStop := FALSE;
    FOR nIdx := 1 TO 4 DO
        GVL_IO.aSimLimitPlus[nIdx] := FALSE;
        GVL_IO.aSimLimitMinus[nIdx] := FALSE;
        GVL_IO.aSimFault[nIdx] := FALSE;
    END_FOR
    IF nStep <> 0 THEN
        (* Test beendet oder abgebrochen: CNC-Stub einmalig zuruecknehmen *)
        GVL_Machine.bCncProgramActive := FALSE; GVL_Machine.bCncMStrobe := FALSE; GVL_Machine.nCncMCode := 0;
        GVL_Machine.rCncSpindleRpm := 0.0;
    END_IF
    nStep := 0;
    RETURN;
END_IF

(* Simulierte HMI: Lebenszeichen alle 100 ms. Simulierter Umrichter: Drehzahl erreicht folgt dem Start. *)
tonHb(IN := NOT tonHb.Q, PT := T#100MS);
IF tonHb.Q AND NOT bHbStop THEN GVL_HMI.stCmd.nHeartbeat := GVL_HMI.stCmd.nHeartbeat + 1; END_IF
GVL_IO.bFuAtSpeed := GVL_IO.bSpindleRun;

(* Simulierte Eingaenge: alles in Ordnung, nur das Sicherheitsrelais steuert der Test *)
GVL_IO.bSafetyRelayFeedback := bRelay AND bDoor;   (* offene Tuer laesst auch das Pilz-Relais abfallen *)
GVL_IO.bDoorClosed   := bDoor;
GVL_IO.bAirOk        := TRUE;
GVL_IO.bExtractionOk := TRUE;
GVL_IO.bFuReady      := TRUE;
GVL_IO.bSpindlePtcOk := TRUE;
GVL_IO.bFieldbusOk   := TRUE;

tonStep(IN := NOT bNext, PT := tWait);
bNext := FALSE;

CASE nStep OF
    0:  (* Start *)
        nFails := 0; sFirstFail := ''; bTestDone := FALSE; bRelay := TRUE;
        GVL_HMI.stCmd.eModeRequest := E_OpMode.Hand;
        nStep := 10; tWait := T#1S; bNext := TRUE;

    10: (* T01 Anlauf: Maschine startet gelatcht, nicht frei *)
        IF tonStep.Q THEN
            (* Eingaenge sind jetzt in Ordnung, aber ohne Quittierung darf die Maschine nicht frei sein (EStop oder Stopped) *)
            IF GVL_HMI.stSts.eState = E_MachState.Idle OR GVL_HMI.stSts.eState = E_MachState.Execute OR GVL_HMI.stSts.bDrivesEnabled THEN sMsg := 'T01 Anlauf ohne Quittierung frei'; bFailNow := TRUE; END_IF
            GVL_HMI.stCmd.bAck := TRUE;
            nStep := 20; tWait := T#1S; bNext := TRUE;
        END_IF

    20: (* T02 Quittierung -> Idle, dann Referenzfahrt anfordern *)
        IF tonStep.Q THEN
            IF GVL_HMI.stSts.eState <> E_MachState.Idle THEN sMsg := 'T02 Quittierung fuehrt nicht nach Idle'; bFailNow := TRUE; END_IF
            GVL_HMI.stCmd.bHomeRequest := TRUE;
            nStep := 30; tWait := T#20S; bNext := TRUE;
        END_IF

    30: (* T03 Referenzfahrt aller Gruppen *)
        IF GVL_HMI.stSts.bAllHomed THEN
            nStep := 40; tWait := T#500MS; bNext := TRUE;
        ELSIF tonStep.Q THEN
            sMsg := 'T03 Referenzfahrt: Zeitueberschreitung'; bFailNow := TRUE;
            nStep := 40; tWait := T#500MS; bNext := TRUE;
        END_IF

    40: (* Tippen: Achse waehlen, 300 ms stabil *)
        IF tonStep.Q THEN
            GVL_HMI.stCmd.nJogAxis := 1;
            nStep := 50; tWait := T#300MS; bNext := TRUE;
        END_IF

    50: (* Tippen+ starten *)
        IF tonStep.Q THEN
            GVL_HMI.stCmd.bJogPlus := TRUE;
            nStep := 60; tWait := T#500MS; bNext := TRUE;
        END_IF

    60: (* T04 Tippen+ aktiv, dann loslassen *)
        IF tonStep.Q THEN
            IF NOT GVL_Machine.bCncJogPlus THEN sMsg := 'T04 Tippen+ startet nicht'; bFailNow := TRUE; END_IF
            GVL_HMI.stCmd.bJogPlus := FALSE;
            nStep := 70; tWait := T#300MS; bNext := TRUE;
        END_IF

    70: (* T05 Tippen stoppt beim Loslassen, dann Taste wieder druecken *)
        IF tonStep.Q THEN
            IF GVL_Machine.bCncJogPlus THEN sMsg := 'T05 Tippen stoppt nicht beim Loslassen'; bFailNow := TRUE; END_IF
            GVL_HMI.stCmd.bJogPlus := TRUE;
            nStep := 80; tWait := T#400MS; bNext := TRUE;
        END_IF

    80: (* NOT-HALT bei gehaltener Tippen-Taste *)
        IF tonStep.Q THEN
            bRelay := FALSE;
            nStep := 90; tWait := T#500MS; bNext := TRUE;
        END_IF

    90: (* T07 NOT-HALT erkannt, Tippen aus, Antriebe weg *)
        IF tonStep.Q THEN
            IF GVL_HMI.stSts.eState <> E_MachState.EStop THEN sMsg := 'T07 NOT-HALT nicht erkannt'; bFailNow := TRUE; END_IF
            IF GVL_Machine.bCncJogPlus THEN sMsg := 'T07b Tippen laeuft bei NOT-HALT weiter'; bFailNow := TRUE; END_IF
            IF GVL_HMI.stSts.bDrivesEnabled THEN sMsg := 'T07c Antriebe bleiben bei NOT-HALT frei'; bFailNow := TRUE; END_IF
            bRelay := TRUE;
            nStep := 100; tWait := T#500MS; bNext := TRUE;
        END_IF

    100: (* T08/T06 Sicherheitskreis wieder zu: kein Wiederanlauf, gehaltene Taste startet nichts *)
        IF tonStep.Q THEN
            IF GVL_HMI.stSts.eState <> E_MachState.EStop THEN sMsg := 'T08 NOT-HALT ohne Quittierung verlassen'; bFailNow := TRUE; END_IF
            IF GVL_Machine.bCncJogPlus THEN sMsg := 'T06 Tippen startet nach NOT-HALT von selbst'; bFailNow := TRUE; END_IF
            GVL_HMI.stCmd.bAck := TRUE;
            nStep := 110; tWait := T#1500MS; bNext := TRUE;
        END_IF

    110: (* T09 Quittierung -> Idle, gehaltene Tippen-Taste startet nicht, dann Spindel in Hand *)
        IF tonStep.Q THEN
            IF GVL_HMI.stSts.eState <> E_MachState.Idle THEN sMsg := 'T09 Quittierung nach NOT-HALT fuehrt nicht nach Idle'; bFailNow := TRUE; END_IF
            IF GVL_Machine.bCncJogPlus THEN sMsg := 'T06b Tippen startet nach Quittierung von selbst'; bFailNow := TRUE; END_IF
            GVL_HMI.stCmd.bJogPlus := FALSE;
            GVL_HMI.stCmd.rSpindleSetRpm := 12000.0;
            GVL_HMI.stCmd.bSpindleOn := TRUE;
            nStep := 120; tWait := T#1500MS; bNext := TRUE;
        END_IF

    120: (* T10 Spindel startet in Hand, Spannung passt zur Drehzahl *)
        IF tonStep.Q THEN
            IF NOT GVL_IO.bSpindleRun THEN sMsg := 'T10 Spindel startet nicht (Hand)'; bFailNow := TRUE; END_IF
            IF ABS(GVL_IO.rSpindleVolt - 7.2) > 0.3 THEN sMsg := 'T10b Spindelspannung passt nicht zu 12000 1/min'; bFailNow := TRUE; END_IF
            bRelay := FALSE;
            nStep := 130; tWait := T#400MS; bNext := TRUE;
        END_IF

    130: (* T11 Spindel stoppt bei NOT-HALT *)
        IF tonStep.Q THEN
            IF GVL_IO.bSpindleRun THEN sMsg := 'T11 Spindel laeuft bei NOT-HALT weiter'; bFailNow := TRUE; END_IF
            bRelay := TRUE;
            nStep := 140; tWait := T#500MS; bNext := TRUE;
        END_IF

    140: (* Quittieren, Spindeltaste bleibt gedrueckt *)
        IF tonStep.Q THEN
            GVL_HMI.stCmd.bAck := TRUE;
            nStep := 150; tWait := T#1500MS; bNext := TRUE;
        END_IF

    150: (* T12 kein Selbstanlauf der Spindel nach Quittierung *)
        IF tonStep.Q THEN
            IF GVL_IO.bSpindleRun THEN sMsg := 'T12 Spindel startet nach Quittierung von selbst'; bFailNow := TRUE; END_IF
            GVL_HMI.stCmd.bSpindleOn := FALSE;
            nStep := 160; tWait := T#11S; bNext := TRUE;   (* Auslaufzeit abwarten: Hand-Start waehrend des Auslaufs wird verworfen (G-11) *)
        END_IF

    160: (* Spindel erneut starten (Auslaufzeit abwarten), danach HMI-Verlust *)
        IF tonStep.Q THEN
            GVL_HMI.stCmd.bSpindleOn := TRUE;
            nStep := 170; tWait := T#13S; bNext := TRUE;
        END_IF

    170: (* T13a Spindel laeuft, dann Lebenszeichen der HMI ausfallen lassen *)
        IF tonStep.Q THEN
            IF NOT GVL_IO.bSpindleRun THEN sMsg := 'T13a Spindel startet nach Stillstand nicht'; bFailNow := TRUE; END_IF
            bHbStop := TRUE;
            nStep := 180; tWait := T#1500MS; bNext := TRUE;
        END_IF

    180: (* T13 Spindel stoppt bei HMI-Verlust, Meldung 330 steht *)
        IF tonStep.Q THEN
            IF GVL_IO.bSpindleRun THEN sMsg := 'T13 Spindel laeuft bei HMI-Verlust weiter'; bFailNow := TRUE; END_IF
            IF NOT GVL_HMI.stSts.aAlarms[13].bActive THEN sMsg := 'T13b Meldung 330 (HMI-Verbindung) fehlt'; bFailNow := TRUE; END_IF
            bHbStop := FALSE;
            nStep := 190; tWait := T#1500MS; bNext := TRUE;
        END_IF

    190: (* T14 kein Selbstanlauf der Spindel bei Rueckkehr der HMI *)
        IF tonStep.Q THEN
            IF GVL_IO.bSpindleRun THEN sMsg := 'T14 Spindel startet bei Rueckkehr der HMI von selbst'; bFailNow := TRUE; END_IF
            GVL_HMI.stCmd.bSpindleOn := FALSE;
            nStep := 300; tWait := T#500MS; bNext := TRUE;
        END_IF

    300: (* G-01 Endschalter: Tippen+ an X starten *)
        IF tonStep.Q THEN
            GVL_HMI.stCmd.nJogAxis := 1;
            GVL_HMI.stCmd.bJogPlus := TRUE;
            nStep := 305; tWait := T#500MS; bNext := TRUE;
        END_IF

    305: (* Ausgangslage: Tippen+ laeuft, dann Endschalter Plus an X ausloesen (Antrieb 3) *)
        IF tonStep.Q THEN
            IF NOT GVL_Machine.bCncJogPlus THEN sMsg := 'T15a Tippen+ startet nicht (Ausgangslage Endschalter)'; bFailNow := TRUE; END_IF
            GVL_IO.aSimLimitPlus[3] := TRUE;
            nStep := 310; tWait := T#400MS; bNext := TRUE;
        END_IF

    310: (* T15 Tippen stoppt am Endschalter, Meldung 302 steht *)
        IF tonStep.Q THEN
            IF GVL_Machine.bCncJogPlus THEN sMsg := 'T15 Tippen stoppt nicht am Endschalter'; bFailNow := TRUE; END_IF
            IF NOT GVL_HMI.stSts.aAlarms[10].bActive THEN sMsg := 'T15b Meldung 302 (Endschalter) fehlt'; bFailNow := TRUE; END_IF
            nStep := 320; tWait := T#400MS; bNext := TRUE;
        END_IF

    320: (* T15c Taste noch gehalten: kein erneuter Start. Dann Taste loslassen und in Richtung Endschalter neu druecken *)
        IF tonStep.Q THEN
            IF GVL_Machine.bCncJogPlus THEN sMsg := 'T15c Tippen startet am Endschalter bei gehaltener Taste erneut'; bFailNow := TRUE; END_IF
            GVL_HMI.stCmd.bJogPlus := FALSE;
            nStep := 325; tWait := T#300MS; bNext := TRUE;
        END_IF

    325:
        IF tonStep.Q THEN
            GVL_HMI.stCmd.bJogRapid := TRUE;
            GVL_HMI.stCmd.bJogPlus := TRUE;
            nStep := 330; tWait := T#400MS; bNext := TRUE;
        END_IF

    330: (* T15d Richtung zum Endschalter gesperrt. Dann Freifahren in Gegenrichtung *)
        IF tonStep.Q THEN
            IF GVL_Machine.bCncJogPlus THEN sMsg := 'T15d Tippen in Richtung Endschalter nicht gesperrt'; bFailNow := TRUE; END_IF
            GVL_HMI.stCmd.bJogPlus := FALSE;
            nStep := 335; tWait := T#300MS; bNext := TRUE;
        END_IF

    335:
        IF tonStep.Q THEN
            GVL_HMI.stCmd.bJogMinus := TRUE;
            nStep := 340; tWait := T#400MS; bNext := TRUE;
        END_IF

    340: (* T16 Freifahren Gegenrichtung moeglich, ohne Eilgang, anderer Achse gesperrt *)
        IF tonStep.Q THEN
            IF NOT GVL_Machine.bCncJogMinus THEN sMsg := 'T16 Freifahren in Gegenrichtung nicht moeglich'; bFailNow := TRUE; END_IF
            IF GVL_Machine.bCncJogRapid THEN sMsg := 'T16b Eilgang beim Freifahren'; bFailNow := TRUE; END_IF
            IF NOT GVL_Machine.bCncJogCreep THEN sMsg := 'T16c Schleichgang-Anforderung fehlt'; bFailNow := TRUE; END_IF
            GVL_HMI.stCmd.bJogMinus := FALSE;
            GVL_HMI.stCmd.bJogRapid := FALSE;
            GVL_HMI.stCmd.nJogAxis := 3;
            nStep := 345; tWait := T#300MS; bNext := TRUE;
        END_IF

    345: (* T16d Endschalter an X: Tippen an Z in beide Richtungen gesperrt *)
        IF tonStep.Q THEN
            GVL_HMI.stCmd.bJogPlus := TRUE;
            nStep := 347; tWait := T#400MS; bNext := TRUE;
        END_IF

    347:
        IF tonStep.Q THEN
            IF GVL_Machine.bCncJogPlus THEN sMsg := 'T16d Tippen an unbeteiligter Achse bei Endschalter erlaubt'; bFailNow := TRUE; END_IF
            GVL_HMI.stCmd.bJogPlus := FALSE;
            GVL_HMI.stCmd.nJogAxis := 1;
            GVL_IO.aSimLimitPlus[3] := FALSE;
            nStep := 350; tWait := T#400MS; bNext := TRUE;
        END_IF

    350: (* Endschalter frei, Meldung quittieren *)
        IF tonStep.Q THEN
            GVL_HMI.stCmd.bAck := TRUE;
            nStep := 360; tWait := T#1500MS; bNext := TRUE;
        END_IF

    360: (* T17 Quittierung nach Endschalter fuehrt nach Idle *)
        IF tonStep.Q THEN
            IF GVL_HMI.stSts.eState <> E_MachState.Idle THEN sMsg := 'T17 Quittierung nach Endschalter fuehrt nicht nach Idle'; bFailNow := TRUE; END_IF
            nStep := 398; tWait := T#6S; bNext := TRUE;   (* Spindel-Auslaufzeit abwarten, sonst wird der Wechsel nach Auto abgelehnt *)
        END_IF

    398: (* Betriebsart Auto anfordern *)
        IF tonStep.Q THEN
            GVL_HMI.stCmd.eModeRequest := E_OpMode.Auto;
            nStep := 400; tWait := T#700MS; bNext := TRUE;
        END_IF

    (* ---- Programmbetrieb mit CNC-Stub (solange TF5200 nicht angebunden ist) ---- *)
    400: (* T18 Auto, Programmstart *)
        IF tonStep.Q THEN
            IF GVL_HMI.stSts.eMode <> E_OpMode.Auto THEN sMsg := 'T18a Betriebsart Auto nicht erreicht'; bFailNow := TRUE; END_IF
            GVL_HMI.stCmd.bStart := TRUE;
            nStep := 405; tWait := T#500MS; bNext := TRUE;
        END_IF

    405: (* CNC meldet Programm aktiv, M3 S12000 *)
        IF tonStep.Q THEN
            IF GVL_HMI.stSts.eState <> E_MachState.Execute THEN sMsg := 'T18b Programmstart nicht angenommen'; bFailNow := TRUE; END_IF
            GVL_Machine.bCncProgramActive := TRUE;
            GVL_Machine.rCncSpindleRpm := 12000.0;
            GVL_Machine.nCncMCode := 3;
            GVL_Machine.bCncMStrobe := TRUE;
            nStep := 410; tWait := T#18S; bNext := TRUE;
        END_IF

    410: (* T19 M3 wird erst quittiert, wenn die Spindel laeuft *)
        IF GVL_Machine.bCncMAck AND NOT GVL_IO.bSpindleRun THEN
            sMsg := 'T19a M3 quittiert, obwohl die Spindel nicht laeuft'; bFailNow := TRUE;
            nStep := 415; tWait := T#300MS; bNext := TRUE;
        ELSIF GVL_IO.bSpindleRun AND GVL_Machine.bCncMAck THEN
            nStep := 415; tWait := T#300MS; bNext := TRUE;
        ELSIF tonStep.Q THEN
            sMsg := 'T19 Spindel startet nach M3 nicht'; bFailNow := TRUE;
            nStep := 415; tWait := T#300MS; bNext := TRUE;
        END_IF

    415: (* T19c S-Wert aus der CNC wirkt, dann M-Code zurueckziehen und Halt *)
        IF tonStep.Q THEN
            IF ABS(GVL_IO.rSpindleVolt - 7.2) > 0.3 THEN sMsg := 'T19c S-Wert aus der CNC nicht uebernommen'; bFailNow := TRUE; END_IF
            GVL_Machine.bCncMStrobe := FALSE; GVL_Machine.nCncMCode := 0;
            GVL_HMI.stCmd.bHold := TRUE;
            nStep := 420; tWait := T#800MS; bNext := TRUE;
        END_IF

    420: (* T20 Vorschubhalt: Zustand Held, Anforderung an die CNC als Pegel *)
        IF tonStep.Q THEN
            IF GVL_HMI.stSts.eState <> E_MachState.Held THEN sMsg := 'T20 Halt nicht angenommen'; bFailNow := TRUE; END_IF
            nStep := 425; tWait := T#2S; bNext := TRUE;
        END_IF

    425:
        IF tonStep.Q THEN
            IF NOT GVL_Machine.bCncHoldReq THEN sMsg := 'T20b Vorschubhalt faellt ab (kein Pegel)'; bFailNow := TRUE; END_IF
            GVL_HMI.stCmd.bStart := TRUE;
            nStep := 430; tWait := T#500MS; bNext := TRUE;
        END_IF

    430: (* T20c Fortsetzen, Halt faellt; dann Vakuum per M10 *)
        IF tonStep.Q THEN
            IF GVL_HMI.stSts.eState <> E_MachState.Execute THEN sMsg := 'T20c Fortsetzen nach Halt nicht moeglich'; bFailNow := TRUE; END_IF
            IF GVL_Machine.bCncHoldReq THEN sMsg := 'T20d Halt bleibt nach Fortsetzen stehen'; bFailNow := TRUE; END_IF
            GVL_Machine.nCncMCode := 10; GVL_Machine.bCncMStrobe := TRUE;
            nStep := 435; tWait := T#400MS; bNext := TRUE;
        END_IF

    435: (* T21a Vakuum an, dann Abbruch *)
        IF tonStep.Q THEN
            IF NOT GVL_IO.bVacuumOut THEN sMsg := 'T21a Vakuum (M10) geht nicht an'; bFailNow := TRUE; END_IF
            GVL_Machine.bCncMStrobe := FALSE; GVL_Machine.nCncMCode := 0;
            GVL_HMI.stCmd.bAbort := TRUE;
            nStep := 440; tWait := T#700MS; bNext := TRUE;
        END_IF

    440: (* T21 Abbruch: Spindel aus, Abbruch an die CNC als Pegel, Vakuum bleibt (G-04) *)
        IF tonStep.Q THEN
            IF GVL_IO.bSpindleRun THEN sMsg := 'T21 Spindel laeuft nach Abbruch weiter'; bFailNow := TRUE; END_IF
            IF NOT GVL_Machine.bCncAbortReq THEN sMsg := 'T21b Abbruch an die CNC fehlt'; bFailNow := TRUE; END_IF
            IF NOT GVL_IO.bVacuumOut THEN sMsg := 'T21c Vakuum faellt bei Abbruch ab'; bFailNow := TRUE; END_IF
            GVL_Machine.bCncProgramActive := FALSE;
            nStep := 445; tWait := T#500MS; bNext := TRUE;
        END_IF

    445: (* T21d Abbruch faellt, wenn die CNC steht. Quittieren, dann M11 *)
        IF tonStep.Q THEN
            IF GVL_Machine.bCncAbortReq THEN sMsg := 'T21d Abbruch bleibt nach Programmstopp stehen'; bFailNow := TRUE; END_IF
            GVL_HMI.stCmd.bAck := TRUE;
            nStep := 450; tWait := T#1500MS; bNext := TRUE;
        END_IF

    450: (* M11 schaltet das Vakuum ab, Zustand Idle *)
        IF tonStep.Q THEN
            IF GVL_HMI.stSts.eState <> E_MachState.Idle THEN sMsg := 'T21e Quittierung nach Abbruch fuehrt nicht nach Idle'; bFailNow := TRUE; END_IF
            GVL_Machine.nCncMCode := 11; GVL_Machine.bCncMStrobe := TRUE;
            nStep := 455; tWait := T#400MS; bNext := TRUE;
        END_IF

    455: (* T21f M11 aus, dann Programm neu starten, Vakuum an, NOT-HALT in Execute *)
        IF tonStep.Q THEN
            IF GVL_IO.bVacuumOut THEN sMsg := 'T21f M11 schaltet das Vakuum nicht ab'; bFailNow := TRUE; END_IF
            GVL_Machine.bCncMStrobe := FALSE; GVL_Machine.nCncMCode := 0;
            GVL_HMI.stCmd.bStart := TRUE;
            nStep := 460; tWait := T#500MS; bNext := TRUE;
        END_IF

    460:
        IF tonStep.Q THEN
            IF GVL_HMI.stSts.eState <> E_MachState.Execute THEN sMsg := 'T22a Programmstart nach Abbruch nicht moeglich'; bFailNow := TRUE; END_IF
            GVL_Machine.bCncProgramActive := TRUE;
            GVL_Machine.nCncMCode := 10; GVL_Machine.bCncMStrobe := TRUE;
            nStep := 465; tWait := T#400MS; bNext := TRUE;
        END_IF

    465: (* NOT-HALT in Execute bei aktiver CNC *)
        IF tonStep.Q THEN
            GVL_Machine.bCncMStrobe := FALSE; GVL_Machine.nCncMCode := 0;
            bRelay := FALSE;
            nStep := 470; tWait := T#600MS; bNext := TRUE;
        END_IF

    470: (* T22 EStop, Abbruch an die CNC, Vakuum bleibt (G-04). Sicherheitskreis wieder zu, quittieren: CNC aktiv, EStop bleibt *)
        IF tonStep.Q THEN
            IF GVL_HMI.stSts.eState <> E_MachState.EStop THEN sMsg := 'T22 NOT-HALT in Execute nicht erkannt'; bFailNow := TRUE; END_IF
            IF NOT GVL_Machine.bCncAbortReq THEN sMsg := 'T22b NOT-HALT in Execute: kein Abbruch an die CNC'; bFailNow := TRUE; END_IF
            IF NOT GVL_IO.bVacuumOut THEN sMsg := 'T22c Vakuum faellt bei NOT-HALT ab'; bFailNow := TRUE; END_IF
            bRelay := TRUE;
            nStep := 475; tWait := T#500MS; bNext := TRUE;
        END_IF

    475:
        IF tonStep.Q THEN
            GVL_HMI.stCmd.bAck := TRUE;
            nStep := 480; tWait := T#800MS; bNext := TRUE;
        END_IF

    480: (* T22d EStop bleibt, solange die CNC noch aktiv meldet *)
        IF tonStep.Q THEN
            IF GVL_HMI.stSts.eState <> E_MachState.EStop THEN sMsg := 'T22d EStop verlassen, obwohl die CNC noch aktiv ist'; bFailNow := TRUE; END_IF
            GVL_Machine.bCncProgramActive := FALSE;
            nStep := 485; tWait := T#500MS; bNext := TRUE;
        END_IF

    485:
        IF tonStep.Q THEN
            GVL_HMI.stCmd.bAck := TRUE;
            nStep := 490; tWait := T#1500MS; bNext := TRUE;
        END_IF

    490: (* T22e Quittierung nach CNC-Stopp fuehrt nach Idle; M11 raeumt auf, zurueck in Hand *)
        IF tonStep.Q THEN
            IF GVL_HMI.stSts.eState <> E_MachState.Idle THEN sMsg := 'T22e Quittierung nach CNC-Stopp fuehrt nicht nach Idle'; bFailNow := TRUE; END_IF
            GVL_Machine.nCncMCode := 11; GVL_Machine.bCncMStrobe := TRUE;
            GVL_HMI.stCmd.eModeRequest := E_OpMode.Hand;
            nStep := 495; tWait := T#600MS; bNext := TRUE;
        END_IF

    495:
        IF tonStep.Q THEN
            GVL_Machine.bCncMStrobe := FALSE; GVL_Machine.nCncMCode := 0;
            GVL_Machine.rCncSpindleRpm := 0.0;
            nStep := 500; tWait := T#2S; bNext := TRUE;
        END_IF

    (* ---- Werkzeugwechsel bei offener Tuer ---- *)
    500: (* Auto, Programm starten, M3 *)
        IF tonStep.Q THEN
            GVL_HMI.stCmd.eModeRequest := E_OpMode.Auto;
            nStep := 502; tWait := T#800MS; bNext := TRUE;
        END_IF

    502:
        IF tonStep.Q THEN
            GVL_HMI.stCmd.bStart := TRUE;
            nStep := 505; tWait := T#500MS; bNext := TRUE;
        END_IF

    505:
        IF tonStep.Q THEN
            GVL_Machine.bCncProgramActive := TRUE;
            GVL_Machine.rCncSpindleRpm := 12000.0;
            GVL_Machine.nCncMCode := 3; GVL_Machine.bCncMStrobe := TRUE;
            nStep := 510; tWait := T#18S; bNext := TRUE;
        END_IF

    510: (* warten, bis die Spindel laeuft und M3 quittiert ist, dann M6 *)
        IF (GVL_IO.bSpindleRun AND GVL_Machine.bCncMAck) OR tonStep.Q THEN
            IF NOT GVL_IO.bSpindleRun THEN sMsg := 'T23 Spindel startet vor dem Werkzeugwechsel nicht'; bFailNow := TRUE; END_IF
            GVL_Machine.bCncMStrobe := FALSE; GVL_Machine.nCncMCode := 0;
            nStep := 512; tWait := T#300MS; bNext := TRUE;
        END_IF

    512:
        IF tonStep.Q THEN
            GVL_Machine.nCncMCode := 6; GVL_Machine.bCncMStrobe := TRUE;
            nStep := 514; tWait := T#500MS; bNext := TRUE;
        END_IF

    514: (* T23a M6 loest Werkzeugwechsel aus, Spindel stoppt, Tuer noch nicht frei *)
        IF tonStep.Q THEN
            IF NOT GVL_HMI.stSts.bToolChangeReq THEN sMsg := 'T23a M6 loest keine Werkzeugwechsel-Aufforderung aus'; bFailNow := TRUE; END_IF
            IF GVL_IO.bSpindleRun THEN sMsg := 'T23b Spindel laeuft bei Werkzeugwechsel weiter'; bFailNow := TRUE; END_IF
            IF GVL_HMI.stSts.bToolChangeDoorRelease THEN sMsg := 'T23c Tuerfreigabe vor Spindelstillstand'; bFailNow := TRUE; END_IF
            GVL_Machine.bCncMStrobe := FALSE; GVL_Machine.nCncMCode := 0;
            nStep := 516; tWait := T#12S; bNext := TRUE;
        END_IF

    516: (* T23d Tuerfreigabe bei Stillstand, dann Tuer oeffnen *)
        IF tonStep.Q THEN
            IF NOT GVL_HMI.stSts.bToolChangeDoorRelease THEN sMsg := 'T23d Tuerfreigabe nach Spindelstillstand fehlt'; bFailNow := TRUE; END_IF
            bDoor := FALSE;
            nStep := 518; tWait := T#800MS; bNext := TRUE;
        END_IF

    518: (* T23e Tuer offen beim Wechsel: Programm bleibt gehalten, kein Abbruch *)
        IF tonStep.Q THEN
            IF GVL_HMI.stSts.eState <> E_MachState.Held THEN sMsg := 'T23e Tuer offen beim Werkzeugwechsel bricht das Programm ab'; bFailNow := TRUE; END_IF
            IF GVL_Machine.bCncAbortReq THEN sMsg := 'T23f Abbruch an die CNC bei Tuer-Oeffnen im Werkzeugwechsel'; bFailNow := TRUE; END_IF
            bDoor := TRUE;
            nStep := 520; tWait := T#600MS; bNext := TRUE;
        END_IF

    520: (* Tuer zu, quittieren *)
        IF tonStep.Q THEN
            GVL_HMI.stCmd.bAck := TRUE;
            nStep := 522; tWait := T#1500MS; bNext := TRUE;
        END_IF

    522: (* T23g weiter im Halt, dann Werkzeug gewechselt *)
        IF tonStep.Q THEN
            IF GVL_HMI.stSts.eState <> E_MachState.Held THEN sMsg := 'T23g nach Tuer zu und Quittieren nicht im Halt'; bFailNow := TRUE; END_IF
            GVL_HMI.stCmd.bToolChangeDone := TRUE;
            nStep := 524; tWait := T#600MS; bNext := TRUE;
        END_IF

    524: (* T23h Wechsel beendet, Fortsetzen nur mit Start, Spindel startet nicht von selbst *)
        IF tonStep.Q THEN
            IF GVL_HMI.stSts.bToolChangeReq THEN sMsg := 'T23h Werkzeugwechsel nicht beendet'; bFailNow := TRUE; END_IF
            IF GVL_HMI.stSts.eState <> E_MachState.Held THEN sMsg := 'T23i Programm laeuft ohne Start weiter'; bFailNow := TRUE; END_IF
            GVL_HMI.stCmd.bStart := TRUE;
            nStep := 526; tWait := T#700MS; bNext := TRUE;
        END_IF

    526: (* T23j Fortsetzen, Spindel aus; dann Tuer oeffnen ohne Werkzeugwechsel *)
        IF tonStep.Q THEN
            IF GVL_HMI.stSts.eState <> E_MachState.Execute THEN sMsg := 'T23j Fortsetzen nach Werkzeugwechsel nicht moeglich'; bFailNow := TRUE; END_IF
            IF GVL_IO.bSpindleRun THEN sMsg := 'T23k Spindel startet nach Werkzeugwechsel von selbst'; bFailNow := TRUE; END_IF
            bDoor := FALSE;
            nStep := 528; tWait := T#800MS; bNext := TRUE;
        END_IF

    528: (* T24 Tuer offen im Programm ohne Werkzeugwechsel: NOT-HALT, Abbruch an die CNC *)
        IF tonStep.Q THEN
            IF GVL_HMI.stSts.eState <> E_MachState.EStop THEN sMsg := 'T24 Tuer offen im Programm fuehrt nicht zu NOT-HALT'; bFailNow := TRUE; END_IF
            IF NOT GVL_Machine.bCncAbortReq THEN sMsg := 'T24b Tuer offen im Programm: kein Abbruch an die CNC'; bFailNow := TRUE; END_IF
            bDoor := TRUE;
            GVL_Machine.bCncProgramActive := FALSE;
            nStep := 530; tWait := T#600MS; bNext := TRUE;
        END_IF

    530:
        IF tonStep.Q THEN
            GVL_HMI.stCmd.bAck := TRUE;
            nStep := 532; tWait := T#1000MS; bNext := TRUE;
        END_IF

    532:
        IF tonStep.Q THEN
            GVL_HMI.stCmd.bAck := TRUE;
            nStep := 534; tWait := T#1500MS; bNext := TRUE;
        END_IF

    534: (* zurueck in Hand *)
        IF tonStep.Q THEN
            IF GVL_HMI.stSts.eState <> E_MachState.Idle THEN sMsg := 'T24c Quittierung nach Tuer-NOT-HALT fuehrt nicht nach Idle'; bFailNow := TRUE; END_IF
            GVL_HMI.stCmd.eModeRequest := E_OpMode.Hand;
            GVL_Machine.rCncSpindleRpm := 0.0;
            nStep := 200; tWait := T#600MS; bNext := TRUE;
        END_IF

    200: (* Ende *)
        IF tonStep.Q THEN
            bTestDone := TRUE;
            nStep := 210;
        END_IF

    210: ;
END_CASE

IF bFailNow THEN
    nFails := nFails + 1;
    IF sFirstFail = '' THEN sFirstFail := sMsg; END_IF
    bFailNow := FALSE;
END_IF
END_PROGRAM
